                   //Initialize the used variable values
                   #temp32TempDword1 := 16#1;
                   #temp16IndexAnalog := 16#0;
                   #temp16IndexDigital := 16#0;
                   #temp16IndexBinary := 16#0;
                   #temp16IndexString := 16#0;
                   //Initialize the Procedure Para index and Name index while changing of Procedure and changing of screen selection b/w Prepared and Current procedure
                   IF ((#statLasProcedureCur <> #ProcedureCur) OR (#statLasProcedureReq <> #ProcedureReq) OR (#statLastReqProcedSelected <> #ProcedureParaType.ProcedureReqCurInd)) THEN
                       #ProcedureParaType.IndexAnalog := 16#0;
                       #ProcedureParaType.NameIndexAnalog := 16#0;
                       #ProcedureParaType.IndexDigital := 16#0;
                       #ProcedureParaType.NameIndexDigital := 16#0;
                       #ProcedureParaType.IndexBinary := 16#0;
                       #ProcedureParaType.NameIndexBinary := 16#0;
                       #ProcedureParaType.IndexString := 16#0;
                       #ProcedureParaType.NameIndexString := 16#0;
                   END_IF;
                   IF (((#ProcedureCur <> 16#0) AND NOT #ProcedureParaType.ProcedureReqCurInd) OR ((#ProcedureReq <> 16#0) AND #ProcedureParaType.ProcedureReqCurInd)) THEN
                       //Used/Mapped parameter count with individual parameter type will written from the Tool
                       #statTotalProcedureParameters := #MAPPED_PROCEDURE_ANALOG + #MAPPED_PROCEDURE_DIGITAL + #MAPPED_PROCEDURE_BINARY + #MAPPED_PROCEDURE_STRING - 1;
                       IF ((#statTotalProcedureParameters >= 0) AND (#statTotalProcedureParameters <= #PROCEDURE_PARAMETER_MAX)) THEN
                           FOR #temp16IndexOfDefinition := #PROCEDURE_PARAMETER_MIN TO #statTotalProcedureParameters BY 1 DO
                               // Condition for allow the loop iteration only within the start and end index
                               IF (((#stat16ProcParaEndIndex - #stat16ProcParaStartIndex) - #temp16IndexOfDefinition + #PROCEDURE_PARAMETER_MIN) >= 0) THEN
                                   #statInternalCurProcParameter[#temp16IndexOfDefinition].index := #tempSetup.stepOrder.parameterIndex[#stat16ProcParaStartIndex + #temp16IndexOfDefinition];  // MiS: content of first parameterIndex to first internal index, content of second parameterIndex to second internal index etc.
                                   #temp16Index := #statInternalCurProcParameter[#temp16IndexOfDefinition].index;//Move index info to the local var
                                   #temp16ParameterType := #tempSetup.step.parameterDefinition[#temp16Index].type;  // Get type of current parameter
                                   #temp16IndexMTP := #tempSetup.step.parameterDefinition[#temp16Index].indexMTP;//Get parameter indexMTP(wrapper DB) from the setup DB.
                                   #temp16IndexIO := #tempSetup.step.parameterDefinition[#temp16Index].indexIO;
                                   //Condition TO check parameter types are in the range
                                   IF (#temp16ParameterType >= #TYPE_NONE) AND (#temp16ParameterType <= #TYPE_STRING) THEN
                                       REGION Copy procedure parameters from input
                                           CASE #temp16ParameterType OF
                                                   // If Parameter type = 1(Analog)
                                               #TYPE_ANALOG:
                                                   REGION Analog
                                                       //Bit Masking funtionality for calculate the used Analog parameter and Position of the Parameter name in the HMI Text List                                              
                                                       #ProcedureParaType.IndexAnalog := #ProcedureParaType.IndexAnalog OR SHL(IN := #temp32TempDword1, N := INT_TO_UINT(#temp16IndexOfDefinition));
                                                       #ProcedureParaType.NameIndexAnalog := #ProcedureParaType.NameIndexAnalog OR SHL(IN := #temp32TempDword1, N := INT_TO_UINT(#temp16Index));
                                                       //WinCC Parameter View Faceplate logic
                                                       //#StatConfigPara.Analog[#temp16IndexIO] := #MTPConfigurationParameterAnalog[#temp16IndexMTP];
                                                       #ProcedureAna[#temp16IndexAnalog].WQC := #ProcedureParameterAnalog[#temp16IndexMTP].WQC;
                                                       #ProcedureAna[#temp16IndexAnalog].ApplyEn := #ProcedureParameterAnalog[#temp16IndexMTP].ApplyEn;
                                                       #ProcedureAna[#temp16IndexAnalog].ApplyInt := #ProcedureParameterAnalog[#temp16IndexMTP].ApplyInt;
                                                       #ProcedureAna[#temp16IndexAnalog].StateChannel := #ProcedureParameterAnalog[#temp16IndexMTP].StateChannel;
                                                       #ProcedureAna[#temp16IndexAnalog].StateOffAut := #ProcedureParameterAnalog[#temp16IndexMTP].StateOffAut;
                                                       #ProcedureAna[#temp16IndexAnalog].StateOpAut := #ProcedureParameterAnalog[#temp16IndexMTP].StateOpAut;
                                                       #ProcedureAna[#temp16IndexAnalog].StateAutAut := #ProcedureParameterAnalog[#temp16IndexMTP].StateAutAut;
                                                       #ProcedureAna[#temp16IndexAnalog].StateOffAct := #ProcedureParameterAnalog[#temp16IndexMTP].StateOffAct;
                                                       #ProcedureAna[#temp16IndexAnalog].StateOpAct := #ProcedureParameterAnalog[#temp16IndexMTP].StateOpAct;
                                                       #ProcedureAna[#temp16IndexAnalog].StateAutAct := #ProcedureParameterAnalog[#temp16IndexMTP].StateAutAct;
                                                       #ProcedureAna[#temp16IndexAnalog].SrcChannel := #ProcedureParameterAnalog[#temp16IndexMTP].SrcChannel;
                                                       #ProcedureAna[#temp16IndexAnalog].SrcExtAut := #ProcedureParameterAnalog[#temp16IndexMTP].SrcExtAut;
                                                       #ProcedureAna[#temp16IndexAnalog].SrcIntAut := #ProcedureParameterAnalog[#temp16IndexMTP].SrcIntAut;
                                                       #ProcedureAna[#temp16IndexAnalog].SrcIntAct := #ProcedureParameterAnalog[#temp16IndexMTP].SrcIntAct;
                                                       #ProcedureAna[#temp16IndexAnalog].SrcExtAct := #ProcedureParameterAnalog[#temp16IndexMTP].SrcExtAct;
                                                       #ProcedureAna[#temp16IndexAnalog].VInt := #ProcedureParameterAnalog[#temp16IndexMTP].VInt;
                                                       #ProcedureAna[#temp16IndexAnalog].VReq := #ProcedureParameterAnalog[#temp16IndexMTP].VReq;
                                                       #ProcedureAna[#temp16IndexAnalog].VOut := #ProcedureParameterAnalog[#temp16IndexMTP].VOut;
                                                       #ProcedureAna[#temp16IndexAnalog].VFbk := #ProcedureParameterAnalog[#temp16IndexMTP].VFbk;
                                                       #ProcedureAna[#temp16IndexAnalog].VSclMin := #ProcedureParameterAnalog[#temp16IndexMTP].VSclMin;
                                                       #ProcedureAna[#temp16IndexAnalog].VSclMax := #ProcedureParameterAnalog[#temp16IndexMTP].VSclMax;
                                                       #ProcedureAna[#temp16IndexAnalog].VUnit := #ProcedureParameterAnalog[#temp16IndexMTP].VUnit;
                                                       #ProcedureAna[#temp16IndexAnalog].VMin := #ProcedureParameterAnalog[#temp16IndexMTP].VMin;
                                                       #ProcedureAna[#temp16IndexAnalog].VMax := #ProcedureParameterAnalog[#temp16IndexMTP].VMax;
                                                       //Write values from WinCC
                                                       IF #ProcedureParameterAnalog[#temp16IndexMTP].OSLevel = #StatProcedureAnalog[#temp16IndexAnalog].OSLevel THEN
                                                           #ProcedureParameterAnalog[#temp16IndexMTP].OSLevel := #ProcedureAna[#temp16IndexAnalog].OSLevel;
                                                       ELSE
                                                           #ProcedureAna[#temp16IndexAnalog].OSLevel := #ProcedureParameterAnalog[#temp16IndexMTP].OSLevel;
                                                       END_IF;
                                                       IF #ProcedureParameterAnalog[#temp16IndexMTP].ApplyExt = #StatProcedureAnalog[#temp16IndexAnalog].ApplyExt THEN
                                                           #ProcedureParameterAnalog[#temp16IndexMTP].ApplyExt := #ProcedureAna[#temp16IndexAnalog].ApplyExt;
                                                       ELSE
                                                           #ProcedureAna[#temp16IndexAnalog].ApplyExt := #ProcedureParameterAnalog[#temp16IndexMTP].ApplyExt;
                                                       END_IF;
                                                       IF #ProcedureParameterAnalog[#temp16IndexMTP].ApplyOp = #StatProcedureAnalog[#temp16IndexAnalog].ApplyOp THEN
                                                           #ProcedureParameterAnalog[#temp16IndexMTP].ApplyOp := #ProcedureAna[#temp16IndexAnalog].ApplyOp;
                                                       ELSE
                                                           #ProcedureAna[#temp16IndexAnalog].ApplyOp := #ProcedureParameterAnalog[#temp16IndexMTP].ApplyOp;
                                                       END_IF;
                                                       IF #ProcedureParameterAnalog[#temp16IndexMTP].Sync = #StatProcedureAnalog[#temp16IndexAnalog].Sync THEN
                                                           #ProcedureParameterAnalog[#temp16IndexMTP].Sync := #ProcedureAna[#temp16IndexAnalog].Sync;
                                                       ELSE
                                                           #ProcedureAna[#temp16IndexAnalog].Sync := #ProcedureParameterAnalog[#temp16IndexMTP].Sync;
                                                       END_IF;
                                                       IF #ProcedureParameterAnalog[#temp16IndexMTP].StateOffOp = #StatProcedureAnalog[#temp16IndexAnalog].StateOffOp THEN
                                                           #ProcedureParameterAnalog[#temp16IndexMTP].StateOffOp := #ProcedureAna[#temp16IndexAnalog].StateOffOp;
                                                       ELSE
                                                           #ProcedureAna[#temp16IndexAnalog].StateOffOp := #ProcedureParameterAnalog[#temp16IndexMTP].StateOffOp;
                                                       END_IF;
                                                       IF #ProcedureParameterAnalog[#temp16IndexMTP].StateOpOp = #StatProcedureAnalog[#temp16IndexAnalog].StateOpOp THEN
                                                           #ProcedureParameterAnalog[#temp16IndexMTP].StateOpOp := #ProcedureAna[#temp16IndexAnalog].StateOpOp;
                                                       ELSE
                                                           #ProcedureAna[#temp16IndexAnalog].StateOpOp := #ProcedureParameterAnalog[#temp16IndexMTP].StateOpOp;
                                                       END_IF;
                                                       IF #ProcedureParameterAnalog[#temp16IndexMTP].StateAutOp = #StatProcedureAnalog[#temp16IndexAnalog].StateAutOp THEN
                                                           #ProcedureParameterAnalog[#temp16IndexMTP].StateAutOp := #ProcedureAna[#temp16IndexAnalog].StateAutOp;
                                                       ELSE
                                                           #ProcedureAna[#temp16IndexAnalog].StateAutOp := #ProcedureParameterAnalog[#temp16IndexMTP].StateAutOp;
                                                       END_IF;
                                                       IF #ProcedureParameterAnalog[#temp16IndexMTP].SrcIntOp = #StatProcedureAnalog[#temp16IndexAnalog].SrcIntOp THEN
                                                           #ProcedureParameterAnalog[#temp16IndexMTP].SrcIntOp := #ProcedureAna[#temp16IndexAnalog].SrcIntOp;
                                                       ELSE
                                                           #ProcedureAna[#temp16IndexAnalog].SrcIntOp := #ProcedureParameterAnalog[#temp16IndexMTP].SrcIntOp;
                                                       END_IF;
                                                       IF #ProcedureParameterAnalog[#temp16IndexMTP].SrcExtOp = #StatProcedureAnalog[#temp16IndexAnalog].SrcExtOp THEN
                                                           #ProcedureParameterAnalog[#temp16IndexMTP].SrcExtOp := #ProcedureAna[#temp16IndexAnalog].SrcExtOp;
                                                       ELSE
                                                           #ProcedureAna[#temp16IndexAnalog].SrcExtOp := #ProcedureParameterAnalog[#temp16IndexMTP].SrcExtOp;
                                                       END_IF;
                                                       IF #ProcedureParameterAnalog[#temp16IndexMTP].VExt = #StatProcedureAnalog[#temp16IndexAnalog].VExt THEN
                                                           #ProcedureParameterAnalog[#temp16IndexMTP].VExt := #ProcedureAna[#temp16IndexAnalog].VExt;
                                                       ELSE
                                                           #ProcedureAna[#temp16IndexAnalog].VExt := #ProcedureParameterAnalog[#temp16IndexMTP].VExt;
                                                       END_IF;
                                                       IF #ProcedureParameterAnalog[#temp16IndexMTP].VOp = #StatProcedureAnalog[#temp16IndexAnalog].VOp THEN
                                                           #ProcedureParameterAnalog[#temp16IndexMTP].VOp := #ProcedureAna[#temp16IndexAnalog].VOp;
                                                       ELSE
                                                           #ProcedureAna[#temp16IndexAnalog].VOp := #ProcedureParameterAnalog[#temp16IndexMTP].VOp;
                                                       END_IF;

                                                       #StatProcedureAnalog[#temp16IndexAnalog].OSLevel := #ProcedureAna[#temp16IndexAnalog].OSLevel;
                                                       #StatProcedureAnalog[#temp16IndexAnalog].ApplyExt := #ProcedureAna[#temp16IndexAnalog].ApplyExt;
                                                       #StatProcedureAnalog[#temp16IndexAnalog].ApplyOp := #ProcedureAna[#temp16IndexAnalog].ApplyOp;
                                                       #StatProcedureAnalog[#temp16IndexAnalog].Sync := #ProcedureAna[#temp16IndexAnalog].Sync;
                                                       #StatProcedureAnalog[#temp16IndexAnalog].StateOffOp := #ProcedureAna[#temp16IndexAnalog].StateOffOp;
                                                       #StatProcedureAnalog[#temp16IndexAnalog].StateOpOp := #ProcedureAna[#temp16IndexAnalog].StateOpOp;
                                                       #StatProcedureAnalog[#temp16IndexAnalog].StateAutOp := #ProcedureAna[#temp16IndexAnalog].StateAutOp;
                                                       #StatProcedureAnalog[#temp16IndexAnalog].SrcIntOp := #ProcedureAna[#temp16IndexAnalog].SrcIntOp;
                                                       #StatProcedureAnalog[#temp16IndexAnalog].SrcExtOp := #ProcedureAna[#temp16IndexAnalog].SrcExtOp;
                                                       #StatProcedureAnalog[#temp16IndexAnalog].VExt := #ProcedureAna[#temp16IndexAnalog].VExt;
                                                       #StatProcedureAnalog[#temp16IndexAnalog].VOp := #ProcedureAna[#temp16IndexAnalog].VOp;

                                                       #temp16IndexAnalog := #temp16IndexAnalog + 1;
                                                   END_REGION
                                                   // If Parameter type = 2(Digital)     
                                               #TYPE_DIGITAL:
                                                   REGION Digital
                                                       //Bit Masking funtionality for calculate the used Digital parameter and Position of the Parameter name in the HMI Text List  
                                                       #ProcedureParaType.IndexDigital := #ProcedureParaType.IndexDigital OR SHL(IN := #temp32TempDword1, N := INT_TO_UINT(#temp16IndexOfDefinition));
                                                       #ProcedureParaType.NameIndexDigital := #ProcedureParaType.NameIndexDigital OR SHL(IN := #temp32TempDword1, N := INT_TO_UINT(#temp16Index));
                                                       //WinCC Parameter View Faceplate logic
                                                       //#StatConfigPara.Digital[#temp16IndexIO] := #MTPConfigurationParameterAnalog[#temp16IndexMTP];
                                                       #ProcedureDint[#temp16IndexDigital].WQC := #ProcedureParameterDigital[#temp16IndexMTP].WQC;
                                                       #ProcedureDint[#temp16IndexDigital].ApplyEn := #ProcedureParameterDigital[#temp16IndexMTP].ApplyEn;
                                                       #ProcedureDint[#temp16IndexDigital].ApplyInt := #ProcedureParameterDigital[#temp16IndexMTP].ApplyInt;
                                                       #ProcedureDint[#temp16IndexDigital].StateChannel := #ProcedureParameterDigital[#temp16IndexMTP].StateChannel;
                                                       #ProcedureDint[#temp16IndexDigital].StateOffAut := #ProcedureParameterDigital[#temp16IndexMTP].StateOffAut;
                                                       #ProcedureDint[#temp16IndexDigital].StateOpAut := #ProcedureParameterDigital[#temp16IndexMTP].StateOpAut;
                                                       #ProcedureDint[#temp16IndexDigital].StateAutAut := #ProcedureParameterDigital[#temp16IndexMTP].StateAutAut;
                                                       #ProcedureDint[#temp16IndexDigital].StateOffAct := #ProcedureParameterDigital[#temp16IndexMTP].StateOffAct;
                                                       #ProcedureDint[#temp16IndexDigital].StateOpAct := #ProcedureParameterDigital[#temp16IndexMTP].StateOpAct;
                                                       #ProcedureDint[#temp16IndexDigital].StateAutAct := #ProcedureParameterDigital[#temp16IndexMTP].StateAutAct;
                                                       #ProcedureDint[#temp16IndexDigital].SrcChannel := #ProcedureParameterDigital[#temp16IndexMTP].SrcChannel;
                                                       #ProcedureDint[#temp16IndexDigital].SrcExtAut := #ProcedureParameterDigital[#temp16IndexMTP].SrcExtAut;
                                                       #ProcedureDint[#temp16IndexDigital].SrcIntAut := #ProcedureParameterDigital[#temp16IndexMTP].SrcIntAut;
                                                       #ProcedureDint[#temp16IndexDigital].SrcIntAct := #ProcedureParameterDigital[#temp16IndexMTP].SrcIntAct;
                                                       #ProcedureDint[#temp16IndexDigital].SrcExtAct := #ProcedureParameterDigital[#temp16IndexMTP].SrcExtAct;
                                                       #ProcedureDint[#temp16IndexDigital].VInt := #ProcedureParameterDigital[#temp16IndexMTP].VInt;
                                                       #ProcedureDint[#temp16IndexDigital].VReq := #ProcedureParameterDigital[#temp16IndexMTP].VReq;
                                                       #ProcedureDint[#temp16IndexDigital].VOut := #ProcedureParameterDigital[#temp16IndexMTP].VOut;
                                                       #ProcedureDint[#temp16IndexDigital].VFbk := #ProcedureParameterDigital[#temp16IndexMTP].VFbk;
                                                       #ProcedureDint[#temp16IndexDigital].VSclMin := #ProcedureParameterDigital[#temp16IndexMTP].VSclMin;
                                                       #ProcedureDint[#temp16IndexDigital].VSclMax := #ProcedureParameterDigital[#temp16IndexMTP].VSclMax;
                                                       #ProcedureDint[#temp16IndexDigital].VUnit := #ProcedureParameterDigital[#temp16IndexMTP].VUnit;
                                                       #ProcedureDint[#temp16IndexDigital].VMin := #ProcedureParameterDigital[#temp16IndexMTP].VMin;
                                                       #ProcedureDint[#temp16IndexDigital].VMax := #ProcedureParameterDigital[#temp16IndexMTP].VMax;
                                                       //Write values from WinCC
                                                       IF #ProcedureParameterDigital[#temp16IndexMTP].OSLevel = #StatProcedureDigital[#temp16IndexDigital].OSLevel THEN
                                                           #ProcedureParameterDigital[#temp16IndexMTP].OSLevel := #ProcedureDint[#temp16IndexDigital].OSLevel;
                                                       ELSE
                                                           #ProcedureDint[#temp16IndexDigital].OSLevel := #ProcedureParameterDigital[#temp16IndexMTP].OSLevel;
                                                       END_IF;
                                                       IF #ProcedureParameterDigital[#temp16IndexMTP].ApplyExt = #StatProcedureDigital[#temp16IndexDigital].ApplyExt THEN
                                                           #ProcedureParameterDigital[#temp16IndexMTP].ApplyExt := #ProcedureDint[#temp16IndexDigital].ApplyExt;
                                                       ELSE
                                                           #ProcedureDint[#temp16IndexDigital].ApplyExt := #ProcedureParameterDigital[#temp16IndexMTP].ApplyExt;
                                                       END_IF;
                                                       IF #ProcedureParameterDigital[#temp16IndexMTP].ApplyOp = #StatProcedureDigital[#temp16IndexDigital].ApplyOp THEN
                                                           #ProcedureParameterDigital[#temp16IndexMTP].ApplyOp := #ProcedureDint[#temp16IndexDigital].ApplyOp;
                                                       ELSE
                                                           #ProcedureDint[#temp16IndexDigital].ApplyOp := #ProcedureParameterDigital[#temp16IndexMTP].ApplyOp;
                                                       END_IF;
                                                       IF #ProcedureParameterDigital[#temp16IndexMTP].Sync = #StatProcedureDigital[#temp16IndexDigital].Sync THEN
                                                           #ProcedureParameterDigital[#temp16IndexMTP].Sync := #ProcedureDint[#temp16IndexDigital].Sync;
                                                       ELSE
                                                           #ProcedureDint[#temp16IndexDigital].Sync := #ProcedureParameterDigital[#temp16IndexMTP].Sync;
                                                       END_IF;
                                                       IF #ProcedureParameterDigital[#temp16IndexMTP].StateOffOp = #StatProcedureDigital[#temp16IndexDigital].StateOffOp THEN
                                                           #ProcedureParameterDigital[#temp16IndexMTP].StateOffOp := #ProcedureDint[#temp16IndexDigital].StateOffOp;
                                                       ELSE
                                                           #ProcedureDint[#temp16IndexDigital].StateOffOp := #ProcedureParameterDigital[#temp16IndexMTP].StateOffOp;
                                                       END_IF;
                                                       IF #ProcedureParameterDigital[#temp16IndexMTP].StateOpOp = #StatProcedureDigital[#temp16IndexDigital].StateOpOp THEN
                                                           #ProcedureParameterDigital[#temp16IndexMTP].StateOpOp := #ProcedureDint[#temp16IndexDigital].StateOpOp;
                                                       ELSE
                                                           #ProcedureDint[#temp16IndexDigital].StateOpOp := #ProcedureParameterDigital[#temp16IndexMTP].StateOpOp;
                                                       END_IF;
                                                       IF #ProcedureParameterDigital[#temp16IndexMTP].StateAutOp = #StatProcedureDigital[#temp16IndexDigital].StateAutOp THEN
                                                           #ProcedureParameterDigital[#temp16IndexMTP].StateAutOp := #ProcedureDint[#temp16IndexDigital].StateAutOp;
                                                       ELSE
                                                           #ProcedureDint[#temp16IndexDigital].StateAutOp := #ProcedureParameterDigital[#temp16IndexMTP].StateAutOp;
                                                       END_IF;
                                                       IF #ProcedureParameterDigital[#temp16IndexMTP].SrcIntOp = #StatProcedureDigital[#temp16IndexDigital].SrcIntOp THEN
                                                           #ProcedureParameterDigital[#temp16IndexMTP].SrcIntOp := #ProcedureDint[#temp16IndexDigital].SrcIntOp;
                                                       ELSE
                                                           #ProcedureDint[#temp16IndexDigital].SrcIntOp := #ProcedureParameterDigital[#temp16IndexMTP].SrcIntOp;
                                                       END_IF;
                                                       IF #ProcedureParameterDigital[#temp16IndexMTP].SrcExtOp = #StatProcedureDigital[#temp16IndexDigital].SrcExtOp THEN
                                                           #ProcedureParameterDigital[#temp16IndexMTP].SrcExtOp := #ProcedureDint[#temp16IndexDigital].SrcExtOp;
                                                       ELSE
                                                           #ProcedureDint[#temp16IndexDigital].SrcExtOp := #ProcedureParameterDigital[#temp16IndexMTP].SrcExtOp;
                                                       END_IF;
                                                       IF #ProcedureParameterDigital[#temp16IndexMTP].VExt = #StatProcedureDigital[#temp16IndexDigital].VExt THEN
                                                           #ProcedureParameterDigital[#temp16IndexMTP].VExt := #ProcedureDint[#temp16IndexDigital].VExt;
                                                       ELSE
                                                           #ProcedureDint[#temp16IndexDigital].VExt := #ProcedureParameterDigital[#temp16IndexMTP].VExt;
                                                       END_IF;
                                                       IF #ProcedureParameterDigital[#temp16IndexMTP].VOp = #StatProcedureDigital[#temp16IndexDigital].VOp THEN
                                                           #ProcedureParameterDigital[#temp16IndexMTP].VOp := #ProcedureDint[#temp16IndexDigital].VOp;
                                                       ELSE
                                                           #ProcedureDint[#temp16IndexDigital].VOp := #ProcedureParameterDigital[#temp16IndexMTP].VOp;
                                                       END_IF;

                                                       #StatProcedureDigital[#temp16IndexDigital].OSLevel := #ProcedureDint[#temp16IndexDigital].OSLevel;
                                                       #StatProcedureDigital[#temp16IndexDigital].ApplyExt := #ProcedureDint[#temp16IndexDigital].ApplyExt;
                                                       #StatProcedureDigital[#temp16IndexDigital].ApplyOp := #ProcedureDint[#temp16IndexDigital].ApplyOp;
                                                       #StatProcedureDigital[#temp16IndexDigital].Sync := #ProcedureDint[#temp16IndexDigital].Sync;
                                                       #StatProcedureDigital[#temp16IndexDigital].StateOffOp := #ProcedureDint[#temp16IndexDigital].StateOffOp;
                                                       #StatProcedureDigital[#temp16IndexDigital].StateOpOp := #ProcedureDint[#temp16IndexDigital].StateOpOp;
                                                       #StatProcedureDigital[#temp16IndexDigital].StateAutOp := #ProcedureDint[#temp16IndexDigital].StateAutOp;
                                                       #StatProcedureDigital[#temp16IndexDigital].SrcIntOp := #ProcedureDint[#temp16IndexDigital].SrcIntOp;
                                                       #StatProcedureDigital[#temp16IndexDigital].SrcExtOp := #ProcedureDint[#temp16IndexDigital].SrcExtOp;
                                                       #StatProcedureDigital[#temp16IndexDigital].VExt := #ProcedureDint[#temp16IndexDigital].VExt;
                                                       #StatProcedureDigital[#temp16IndexDigital].VOp := #ProcedureDint[#temp16IndexDigital].VOp;

                                                       #temp16IndexDigital := #temp16IndexDigital + 1;
                                                   END_REGION
                                                   // If Parameter type = 3(Binary)    
                                               #TYPE_BINARY:
                                                   REGION Binary
                                                       //Bit Masking funtionality for calculate the used Binary parameter and Position of the Parameter name in the HMI Text List  
                                                       #ProcedureParaType.IndexBinary := #ProcedureParaType.IndexBinary OR SHL(IN := #temp32TempDword1, N := INT_TO_UINT(#temp16IndexOfDefinition));
                                                       #ProcedureParaType.NameIndexBinary := #ProcedureParaType.NameIndexBinary OR SHL(IN := #temp32TempDword1, N := INT_TO_UINT(#temp16Index));
                                                       //WinCC Parameter View Faceplate logic
                                                       //#StatConfigPara.Binary[#temp16IndexIO] := #MTPConfigurationParameterAnalog[#temp16IndexMTP];
                                                       #ProcedureBin[#temp16IndexBinary].WQC := #ProcedureParameterBinary[#temp16IndexMTP].WQC;
                                                       #ProcedureBin[#temp16IndexBinary].ApplyEn := #ProcedureParameterBinary[#temp16IndexMTP].ApplyEn;
                                                       #ProcedureBin[#temp16IndexBinary].ApplyInt := #ProcedureParameterBinary[#temp16IndexMTP].ApplyInt;
                                                       #ProcedureBin[#temp16IndexBinary].StateChannel := #ProcedureParameterBinary[#temp16IndexMTP].StateChannel;
                                                       #ProcedureBin[#temp16IndexBinary].StateOffAut := #ProcedureParameterBinary[#temp16IndexMTP].StateOffAut;
                                                       #ProcedureBin[#temp16IndexBinary].StateOpAut := #ProcedureParameterBinary[#temp16IndexMTP].StateOpAut;
                                                       #ProcedureBin[#temp16IndexBinary].StateAutAut := #ProcedureParameterBinary[#temp16IndexMTP].StateAutAut;
                                                       #ProcedureBin[#temp16IndexBinary].StateOffAct := #ProcedureParameterBinary[#temp16IndexMTP].StateOffAct;
                                                       #ProcedureBin[#temp16IndexBinary].StateOpAct := #ProcedureParameterBinary[#temp16IndexMTP].StateOpAct;
                                                       #ProcedureBin[#temp16IndexBinary].StateAutAct := #ProcedureParameterBinary[#temp16IndexMTP].StateAutAct;
                                                       #ProcedureBin[#temp16IndexBinary].SrcChannel := #ProcedureParameterBinary[#temp16IndexMTP].SrcChannel;
                                                       #ProcedureBin[#temp16IndexBinary].SrcExtAut := #ProcedureParameterBinary[#temp16IndexMTP].SrcExtAut;
                                                       #ProcedureBin[#temp16IndexBinary].SrcIntAut := #ProcedureParameterBinary[#temp16IndexMTP].SrcIntAut;
                                                       #ProcedureBin[#temp16IndexBinary].SrcIntAct := #ProcedureParameterBinary[#temp16IndexMTP].SrcIntAct;
                                                       #ProcedureBin[#temp16IndexBinary].SrcExtAct := #ProcedureParameterBinary[#temp16IndexMTP].SrcExtAct;
                                                       #ProcedureBin[#temp16IndexBinary].VInt := #ProcedureParameterBinary[#temp16IndexMTP].VInt;
                                                       #ProcedureBin[#temp16IndexBinary].VReq := #ProcedureParameterBinary[#temp16IndexMTP].VReq;
                                                       #ProcedureBin[#temp16IndexBinary].VOut := #ProcedureParameterBinary[#temp16IndexMTP].VOut;
                                                       #ProcedureBin[#temp16IndexBinary].VFbk := #ProcedureParameterBinary[#temp16IndexMTP].VFbk;

                                                       //Write values from WinCC
                                                       IF #ProcedureParameterBinary[#temp16IndexMTP].OSLevel = #StatProcedureBinary[#temp16IndexBinary].OSLevel THEN
                                                           #ProcedureParameterBinary[#temp16IndexMTP].OSLevel := #ProcedureBin[#temp16IndexBinary].OSLevel;
                                                       ELSE
                                                           #ProcedureBin[#temp16IndexBinary].OSLevel := #ProcedureParameterBinary[#temp16IndexMTP].OSLevel;
                                                       END_IF;
                                                       IF #ProcedureParameterBinary[#temp16IndexMTP].ApplyExt = #StatProcedureBinary[#temp16IndexBinary].ApplyExt THEN
                                                           #ProcedureParameterBinary[#temp16IndexMTP].ApplyExt := #ProcedureBin[#temp16IndexBinary].ApplyExt;
                                                       ELSE
                                                           #ProcedureBin[#temp16IndexBinary].ApplyExt := #ProcedureParameterBinary[#temp16IndexMTP].ApplyExt;
                                                       END_IF;
                                                       IF #ProcedureParameterBinary[#temp16IndexMTP].ApplyOp = #StatProcedureBinary[#temp16IndexBinary].ApplyOp THEN
                                                           #ProcedureParameterBinary[#temp16IndexMTP].ApplyOp := #ProcedureBin[#temp16IndexBinary].ApplyOp;
                                                       ELSE
                                                           #ProcedureBin[#temp16IndexBinary].ApplyOp := #ProcedureParameterBinary[#temp16IndexMTP].ApplyOp;
                                                       END_IF;
                                                       IF #ProcedureParameterBinary[#temp16IndexMTP].Sync = #StatProcedureBinary[#temp16IndexBinary].Sync THEN
                                                           #ProcedureParameterBinary[#temp16IndexMTP].Sync := #ProcedureBin[#temp16IndexBinary].Sync;
                                                       ELSE
                                                           #ProcedureBin[#temp16IndexBinary].Sync := #ProcedureParameterBinary[#temp16IndexMTP].Sync;
                                                       END_IF;
                                                       IF #ProcedureParameterBinary[#temp16IndexMTP].StateOffOp = #StatProcedureBinary[#temp16IndexBinary].StateOffOp THEN
                                                           #ProcedureParameterBinary[#temp16IndexMTP].StateOffOp := #ProcedureBin[#temp16IndexBinary].StateOffOp;
                                                       ELSE
                                                           #ProcedureBin[#temp16IndexBinary].StateOffOp := #ProcedureParameterBinary[#temp16IndexMTP].StateOffOp;
                                                       END_IF;
                                                       IF #ProcedureParameterBinary[#temp16IndexMTP].StateOpOp = #StatProcedureBinary[#temp16IndexBinary].StateOpOp THEN
                                                           #ProcedureParameterBinary[#temp16IndexMTP].StateOpOp := #ProcedureBin[#temp16IndexBinary].StateOpOp;
                                                       ELSE
                                                           #ProcedureBin[#temp16IndexBinary].StateOpOp := #ProcedureParameterBinary[#temp16IndexMTP].StateOpOp;
                                                       END_IF;
                                                       IF #ProcedureParameterBinary[#temp16IndexMTP].StateAutOp = #StatProcedureBinary[#temp16IndexBinary].StateAutOp THEN
                                                           #ProcedureParameterBinary[#temp16IndexMTP].StateAutOp := #ProcedureBin[#temp16IndexBinary].StateAutOp;
                                                       ELSE
                                                           #ProcedureBin[#temp16IndexBinary].StateAutOp := #ProcedureParameterBinary[#temp16IndexMTP].StateAutOp;
                                                       END_IF;
                                                       IF #ProcedureParameterBinary[#temp16IndexMTP].SrcIntOp = #StatProcedureBinary[#temp16IndexBinary].SrcIntOp THEN
                                                           #ProcedureParameterBinary[#temp16IndexMTP].SrcIntOp := #ProcedureBin[#temp16IndexBinary].SrcIntOp;
                                                       ELSE
                                                           #ProcedureBin[#temp16IndexBinary].SrcIntOp := #ProcedureParameterBinary[#temp16IndexMTP].SrcIntOp;
                                                       END_IF;
                                                       IF #ProcedureParameterBinary[#temp16IndexMTP].SrcExtOp = #StatProcedureBinary[#temp16IndexBinary].SrcExtOp THEN
                                                           #ProcedureParameterBinary[#temp16IndexMTP].SrcExtOp := #ProcedureBin[#temp16IndexBinary].SrcExtOp;
                                                       ELSE
                                                           #ProcedureBin[#temp16IndexBinary].SrcExtOp := #ProcedureParameterBinary[#temp16IndexMTP].SrcExtOp;
                                                       END_IF;
                                                       IF #ProcedureParameterBinary[#temp16IndexMTP].VExt = #StatProcedureBinary[#temp16IndexBinary].VExt THEN
                                                           #ProcedureParameterBinary[#temp16IndexMTP].VExt := #ProcedureBin[#temp16IndexBinary].VExt;
                                                       ELSE
                                                           #ProcedureBin[#temp16IndexBinary].VExt := #ProcedureParameterBinary[#temp16IndexMTP].VExt;
                                                       END_IF;
                                                       IF #ProcedureParameterBinary[#temp16IndexMTP].VOp = #StatProcedureBinary[#temp16IndexBinary].VOp THEN
                                                           #ProcedureParameterBinary[#temp16IndexMTP].VOp := #ProcedureBin[#temp16IndexBinary].VOp;
                                                       ELSE
                                                           #ProcedureBin[#temp16IndexBinary].VOp := #ProcedureParameterBinary[#temp16IndexMTP].VOp;
                                                       END_IF;

                                                       #StatProcedureBinary[#temp16IndexBinary].OSLevel := #ProcedureBin[#temp16IndexBinary].OSLevel;
                                                       #StatProcedureBinary[#temp16IndexBinary].ApplyExt := #ProcedureBin[#temp16IndexBinary].ApplyExt;
                                                       #StatProcedureBinary[#temp16IndexBinary].ApplyOp := #ProcedureBin[#temp16IndexBinary].ApplyOp;
                                                       #StatProcedureBinary[#temp16IndexBinary].Sync := #ProcedureBin[#temp16IndexBinary].Sync;
                                                       #StatProcedureBinary[#temp16IndexBinary].StateOffOp := #ProcedureBin[#temp16IndexBinary].StateOffOp;
                                                       #StatProcedureBinary[#temp16IndexBinary].StateOpOp := #ProcedureBin[#temp16IndexBinary].StateOpOp;
                                                       #StatProcedureBinary[#temp16IndexBinary].StateAutOp := #ProcedureBin[#temp16IndexBinary].StateAutOp;
                                                       #StatProcedureBinary[#temp16IndexBinary].SrcIntOp := #ProcedureBin[#temp16IndexBinary].SrcIntOp;
                                                       #StatProcedureBinary[#temp16IndexBinary].SrcExtOp := #ProcedureBin[#temp16IndexBinary].SrcExtOp;
                                                       #StatProcedureBinary[#temp16IndexBinary].VExt := #ProcedureBin[#temp16IndexBinary].VExt;
                                                       #StatProcedureBinary[#temp16IndexBinary].VOp := #ProcedureBin[#temp16IndexBinary].VOp;

                                                       #temp16IndexBinary := #temp16IndexBinary + 1;
                                                   END_REGION
                                                   // If Parameter type = 4(String)    
                                               #TYPE_STRING:
                                                   REGION String
                                                       //Bit Masking funtionality for calculate the used String parameter and Position of the Parameter name in the HMI Text List  
                                                       #ProcedureParaType.IndexString := #ProcedureParaType.IndexString OR SHL(IN := #temp32TempDword1, N := INT_TO_UINT(#temp16IndexOfDefinition));
                                                       #ProcedureParaType.NameIndexString := #ProcedureParaType.NameIndexString OR SHL(IN := #temp32TempDword1, N := INT_TO_UINT(#temp16Index));
                                                       //WinCC Parameter View Faceplate logic
                                                       //#StatConfigPara."String"[#temp16IndexIO] := #MTPConfigurationParameterString[#temp16IndexMTP];
                                                       #ProcedureString[#temp16IndexString].WQC := #ProcedureParameterString[#temp16IndexMTP].WQC;
                                                       #ProcedureString[#temp16IndexString].ApplyEn := #ProcedureParameterString[#temp16IndexMTP].ApplyEn;
                                                       #ProcedureString[#temp16IndexString].ApplyInt := #ProcedureParameterString[#temp16IndexMTP].ApplyInt;
                                                       #ProcedureString[#temp16IndexString].StateChannel := #ProcedureParameterString[#temp16IndexMTP].StateChannel;
                                                       #ProcedureString[#temp16IndexString].StateOffAut := #ProcedureParameterString[#temp16IndexMTP].StateOffAut;
                                                       #ProcedureString[#temp16IndexString].StateOpAut := #ProcedureParameterString[#temp16IndexMTP].StateOpAut;
                                                       #ProcedureString[#temp16IndexString].StateAutAut := #ProcedureParameterString[#temp16IndexMTP].StateAutAut;
                                                       #ProcedureString[#temp16IndexString].StateOffAct := #ProcedureParameterString[#temp16IndexMTP].StateOffAct;
                                                       #ProcedureString[#temp16IndexString].StateOpAct := #ProcedureParameterString[#temp16IndexMTP].StateOpAct;
                                                       #ProcedureString[#temp16IndexString].StateAutAct := #ProcedureParameterString[#temp16IndexMTP].StateAutAct;
                                                       #ProcedureString[#temp16IndexString].SrcChannel := #ProcedureParameterString[#temp16IndexMTP].SrcChannel;
                                                       #ProcedureString[#temp16IndexString].SrcExtAut := #ProcedureParameterString[#temp16IndexMTP].SrcExtAut;
                                                       #ProcedureString[#temp16IndexString].SrcIntAut := #ProcedureParameterString[#temp16IndexMTP].SrcIntAut;
                                                       #ProcedureString[#temp16IndexString].SrcIntAct := #ProcedureParameterString[#temp16IndexMTP].SrcIntAct;
                                                       #ProcedureString[#temp16IndexString].SrcExtAct := #ProcedureParameterString[#temp16IndexMTP].SrcExtAct;
                                                       #ProcedureString[#temp16IndexString].VInt := #ProcedureParameterString[#temp16IndexMTP].VInt;
                                                       #ProcedureString[#temp16IndexString].VReq := #ProcedureParameterString[#temp16IndexMTP].VReq;
                                                       #ProcedureString[#temp16IndexString].VOut := #ProcedureParameterString[#temp16IndexMTP].VOut;
                                                       #ProcedureString[#temp16IndexString].VFbk := #ProcedureParameterString[#temp16IndexMTP].VFbk;

                                                       //Write values from WinCC
                                                       IF #ProcedureParameterString[#temp16IndexMTP].OSLevel = #StatProcedureString[#temp16IndexString].OSLevel THEN
                                                           #ProcedureParameterString[#temp16IndexMTP].OSLevel := #ProcedureString[#temp16IndexString].OSLevel;
                                                       ELSE
                                                           #ProcedureString[#temp16IndexString].OSLevel := #ProcedureParameterString[#temp16IndexMTP].OSLevel;
                                                       END_IF;
                                                       IF #ProcedureParameterString[#temp16IndexMTP].ApplyExt = #StatProcedureString[#temp16IndexString].ApplyExt THEN
                                                           #ProcedureParameterString[#temp16IndexMTP].ApplyExt := #ProcedureString[#temp16IndexString].ApplyExt;
                                                       ELSE
                                                           #ProcedureString[#temp16IndexString].ApplyExt := #ProcedureParameterString[#temp16IndexMTP].ApplyExt;
                                                       END_IF;
                                                       IF #ProcedureParameterString[#temp16IndexMTP].ApplyOp = #StatProcedureString[#temp16IndexString].ApplyOp THEN
                                                           #ProcedureParameterString[#temp16IndexMTP].ApplyOp := #ProcedureString[#temp16IndexString].ApplyOp;
                                                       ELSE
                                                           #ProcedureString[#temp16IndexString].ApplyOp := #ProcedureParameterString[#temp16IndexMTP].ApplyOp;
                                                       END_IF;
                                                       IF #ProcedureParameterString[#temp16IndexMTP].Sync = #StatProcedureString[#temp16IndexString].Sync THEN
                                                           #ProcedureParameterString[#temp16IndexMTP].Sync := #ProcedureString[#temp16IndexString].Sync;
                                                       ELSE
                                                           #ProcedureString[#temp16IndexString].Sync := #ProcedureParameterString[#temp16IndexMTP].Sync;
                                                       END_IF;
                                                       IF #ProcedureParameterString[#temp16IndexMTP].StateOffOp = #StatProcedureString[#temp16IndexString].StateOffOp THEN
                                                           #ProcedureParameterString[#temp16IndexMTP].StateOffOp := #ProcedureString[#temp16IndexString].StateOffOp;
                                                       ELSE
                                                           #ProcedureString[#temp16IndexString].StateOffOp := #ProcedureParameterString[#temp16IndexMTP].StateOffOp;
                                                       END_IF;
                                                       IF #ProcedureParameterString[#temp16IndexMTP].StateOpOp = #StatProcedureString[#temp16IndexString].StateOpOp THEN
                                                           #ProcedureParameterString[#temp16IndexMTP].StateOpOp := #ProcedureString[#temp16IndexString].StateOpOp;
                                                       ELSE
                                                           #ProcedureString[#temp16IndexString].StateOpOp := #ProcedureParameterString[#temp16IndexMTP].StateOpOp;
                                                       END_IF;
                                                       IF #ProcedureParameterString[#temp16IndexMTP].StateAutOp = #StatProcedureString[#temp16IndexString].StateAutOp THEN
                                                           #ProcedureParameterString[#temp16IndexMTP].StateAutOp := #ProcedureString[#temp16IndexString].StateAutOp;
                                                       ELSE
                                                           #ProcedureString[#temp16IndexString].StateAutOp := #ProcedureParameterString[#temp16IndexMTP].StateAutOp;
                                                       END_IF;
                                                       IF #ProcedureParameterString[#temp16IndexMTP].SrcIntOp = #StatProcedureString[#temp16IndexString].SrcIntOp THEN
                                                           #ProcedureParameterString[#temp16IndexMTP].SrcIntOp := #ProcedureString[#temp16IndexString].SrcIntOp;
                                                       ELSE
                                                           #ProcedureString[#temp16IndexString].SrcIntOp := #ProcedureParameterString[#temp16IndexMTP].SrcIntOp;
                                                       END_IF;
                                                       IF #ProcedureParameterString[#temp16IndexMTP].SrcExtOp = #StatProcedureString[#temp16IndexString].SrcExtOp THEN
                                                           #ProcedureParameterString[#temp16IndexMTP].SrcExtOp := #ProcedureString[#temp16IndexString].SrcExtOp;
                                                       ELSE
                                                           #ProcedureString[#temp16IndexString].SrcExtOp := #ProcedureParameterString[#temp16IndexMTP].SrcExtOp;
                                                       END_IF;
                                                       IF #ProcedureParameterString[#temp16IndexMTP].VExt = #StatProcedureString[#temp16IndexString].VExt THEN
                                                           #ProcedureParameterString[#temp16IndexMTP].VExt := #ProcedureString[#temp16IndexString].VExt;
                                                       ELSE
                                                           #ProcedureString[#temp16IndexString].VExt := #ProcedureParameterString[#temp16IndexMTP].VExt;
                                                       END_IF;
                                                       IF #ProcedureParameterString[#temp16IndexMTP].VOp = #StatProcedureString[#temp16IndexString].VOp THEN
                                                           #ProcedureParameterString[#temp16IndexMTP].VOp := #ProcedureString[#temp16IndexString].VOp;
                                                       ELSE
                                                           #ProcedureString[#temp16IndexString].VOp := #ProcedureParameterString[#temp16IndexMTP].VOp;
                                                       END_IF;

                                                       #StatProcedureString[#temp16IndexString].OSLevel := #ProcedureString[#temp16IndexString].OSLevel;
                                                       #StatProcedureString[#temp16IndexString].ApplyExt := #ProcedureString[#temp16IndexString].ApplyExt;
                                                       #StatProcedureString[#temp16IndexString].ApplyOp := #ProcedureString[#temp16IndexString].ApplyOp;
                                                       #StatProcedureString[#temp16IndexString].Sync := #ProcedureString[#temp16IndexString].Sync;
                                                       #StatProcedureString[#temp16IndexString].StateOffOp := #ProcedureString[#temp16IndexString].StateOffOp;
                                                       #StatProcedureString[#temp16IndexString].StateOpOp := #ProcedureString[#temp16IndexString].StateOpOp;
                                                       #StatProcedureString[#temp16IndexString].StateAutOp := #ProcedureString[#temp16IndexString].StateAutOp;
                                                       #StatProcedureString[#temp16IndexString].SrcIntOp := #ProcedureString[#temp16IndexString].SrcIntOp;
                                                       #StatProcedureString[#temp16IndexString].SrcExtOp := #ProcedureString[#temp16IndexString].SrcExtOp;
                                                       #StatProcedureString[#temp16IndexString].VExt := #ProcedureString[#temp16IndexString].VExt;
                                                       #StatProcedureString[#temp16IndexString].VOp := #ProcedureString[#temp16IndexString].VOp;

                                                       #temp16IndexString := #temp16IndexString + 1;
                                                   END_REGION
                                           END_CASE;
                                       END_REGION
                                   END_IF;
                               END_IF;
                           END_FOR;
                       END_IF;
                   END_IF;
               END_IF;
           END_REGION
       END_REGION

       REGION Process In Values

           REGION Get Start and End index details of the Current /Prepared procedure
               //Current/Prepared procedure selection for parameter display in the faceplate
               //#stat32PrecedureProcessInMap := -1;
               IF NOT (#ProcessInValueType.ProcedureReqCurInd) THEN
                   #stat32PrecedureProcessInMap := #tempSetup.procedure.procedure[#stat16ProceCurIndex].ProcedureProcessInMap[0];
               ELSIF (#ProcessInValueType.ProcedureReqCurInd) THEN
                   #stat32PrecedureProcessInMap := #tempSetup.procedure.procedure[#stat16ProceReqIndex].ProcedureProcessInMap[0];
               END_IF;
           END_REGION
           //Initialize the used variable values        
           #temp32TempDword1 := 16#1;
           #temp16IndexAnalog := 16#0;
           #temp16IndexDigital := 16#0;
           #temp16IndexBinary := 16#0;
           #temp16IndexString := 16#0;
           //Initialize the Process In Value index and Name index while changing of Procedure and changing of screen selection b/w Prepared and Current procedure
           IF ((#statLasProcedureCur <> #ProcedureCur) OR (#statLasProcedureReq <> #ProcedureReq) OR (#StatLastProceselProcessIn <> #ProcessInValueType.ProcedureReqCurInd)
               OR (((#ProcedureCur = 16#0) AND NOT #ProcessInValueType.ProcedureReqCurInd) OR ((#ProcedureReq = 16#0) AND #ProcessInValueType.ProcedureReqCurInd))) THEN
               #ProcessInValueType.IndexAnalog := 16#0;
               #ProcessInValueType.NameIndexAnalog := 16#0;
               #ProcessInValueType.IndexDigital := 16#0;
               #ProcessInValueType.NameIndexDigital := 16#0;
               #ProcessInValueType.IndexBinary := 16#0;
               #ProcessInValueType.NameIndexBinary := 16#0;
               #ProcessInValueType.IndexString := 16#0;
               #ProcessInValueType.NameIndexString := 16#0;
           END_IF;
           //Used/Mapped parameter count with individual parameter type will written from the Tool
           #statTotalProcessInValues := #MAPPED_PROCESS_IN_ANALOG + #MAPPED_PROCESS_IN_DIGITAL + #MAPPED_PROCESS_IN_BINARY + #MAPPED_PROCESS_IN_STRING - 1;
           IF (((#ProcedureCur <> 16#0) AND NOT #ProcessInValueType.ProcedureReqCurInd) OR ((#ProcedureReq <> 16#0) AND #ProcessInValueType.ProcedureReqCurInd)) THEN
               IF ((#statTotalProcessInValues >= 0) AND (#statTotalProcessInValues <= #PROCESS_VALUES_IN_MAX)) THEN
                   #temp16IndexOfDefinitionProcessIn := 16#0;
                   FOR #temp16IndexOfDefinition := #PROCESS_VALUES_IN_MIN TO #statTotalProcessInValues BY 1 DO
                       #temp16ParameterCMAddress := BYTE_TO_INT(#tempSetup.processValueInData.definition[#temp16IndexOfDefinition].controlModule);
                       #temp16ParameterType := #tempSetup.processValueInData.definition[#temp16IndexOfDefinition].type;
                       #temp16IndexMTP := #tempSetup.processValueInData.definition[#temp16IndexOfDefinition].indexMTP;
                       #tempUsed := #tempSetup.processValueInData.used;
                       // Find the procedure information assigned with the processIn values
                       IF (((#stat32PrecedureProcessInMap AND SHL(IN := #temp32TempDword1, N := INT_TO_UINT(#temp16IndexOfDefinition))) <> 0) = TRUE) THEN
                           #temp16IndexIO := #tempSetup.processValueInData.definition[#temp16IndexOfDefinition].indexIO;

                           IF (#temp16ParameterCMAddress <> 255) AND (#temp16ParameterCMAddress >= #NUMBER_OF_CONTROLMODULES_MIN) AND (#temp16ParameterCMAddress <= #NUMBER_OF_CONTROLMODULES)
                               AND (#temp16ParameterType >= #TYPE_NONE) AND (#temp16ParameterType <= #TYPE_STRING) THEN
                               #temp16TempInt1 := #temp16ParameterCMAddress / 32;    //DWORD - Adress
                               #temp16TempInt2 := #temp16ParameterCMAddress MOD 32;  //Bit - Adress
                               //If parameter is forced (FRC) --> Parameter is used
                               IF (((#tempUsed[#temp16TempInt1] AND SHL(IN := #temp32TempDword1, N := INT_TO_UINT(#temp16TempInt2))) <> 0) = TRUE) THEN
                                   CASE #temp16ParameterType OF
                                           // Check of mode is done in satellite blocks
                                       #TYPE_ANALOG:
                                           REGION Analog
                                               //Bit Masking funtionality for calculate the used Analog parameter and Position of the Parameter name in the HMI Text List 
                                               #ProcessInValueType.IndexAnalog := #ProcessInValueType.IndexAnalog OR SHL(IN := #temp32TempDword1, N := INT_TO_UINT(#temp16IndexOfDefinitionProcessIn));
                                               #ProcessInValueType.NameIndexAnalog := #ProcessInValueType.NameIndexAnalog OR SHL(IN := #temp32TempDword1, N := INT_TO_UINT(#temp16IndexOfDefinition));
                                               IF ((#temp16IndexIO >= #PROCESS_VALUES_IN_MIN) AND (#temp16IndexIO <= #PROCESS_VALUES_IN_ANALOG_MAX)) THEN
                                                   //WinCC Parameter View Faceplate logic
                                                   #ProcessInAna[#temp16IndexAnalog].WQC := #ProcessValueInAnalog[#temp16IndexMTP].WQC;
                                                   #ProcessInAna[#temp16IndexAnalog].OSLevel := #ProcessValueInAnalog[#temp16IndexMTP].OSLevel;
                                                   #ProcessInAna[#temp16IndexAnalog].V := #ProcessValueInAnalog[#temp16IndexMTP].V;
                                                   #ProcessInAna[#temp16IndexAnalog].VQC := #ProcessValueInAnalog[#temp16IndexMTP].VQC;
                                                   #ProcessInAna[#temp16IndexAnalog].SclMinCur := #ProcessValueInAnalog[#temp16IndexMTP].SclMinCur;
                                                   #ProcessInAna[#temp16IndexAnalog].SclMaxCur := #ProcessValueInAnalog[#temp16IndexMTP].SclMaxCur;
                                                   #ProcessInAna[#temp16IndexAnalog].UnitCur := #ProcessValueInAnalog[#temp16IndexMTP].UnitCur;
                                                   #ProcessInAna[#temp16IndexAnalog].SclMinExt := #ProcessValueInAnalog[#temp16IndexMTP].SclMinExt;
                                                   #ProcessInAna[#temp16IndexAnalog].SclMaxExt := #ProcessValueInAnalog[#temp16IndexMTP].SclMaxExt;
                                                   #ProcessInAna[#temp16IndexAnalog].UnitExt := #ProcessValueInAnalog[#temp16IndexMTP].UnitExt;
                                                   #ProcessInAna[#temp16IndexAnalog].Apply := #ProcessValueInAnalog[#temp16IndexMTP].Apply;
                                                   #ProcessInAna[#temp16IndexAnalog].ApplyEn := #ProcessValueInAnalog[#temp16IndexMTP].ApplyEn;
                                               END_IF;
                                               #temp16IndexAnalog := #temp16IndexAnalog + 1;
                                           END_REGION
                                       #TYPE_DIGITAL:
                                           REGION Digital
                                               //Bit Masking funtionality for calculate the used Digital parameter and Position of the Parameter name in the HMI Text List 
                                               #ProcessInValueType.IndexDigital := #ProcessInValueType.IndexDigital OR SHL(IN := #temp32TempDword1, N := INT_TO_UINT(#temp16IndexOfDefinitionProcessIn));
                                               #ProcessInValueType.NameIndexDigital := #ProcessInValueType.NameIndexDigital OR SHL(IN := #temp32TempDword1, N := INT_TO_UINT(#temp16IndexOfDefinition));
                                               IF ((#temp16IndexIO >= #PROCESS_VALUES_IN_MIN) AND (#temp16IndexIO <= #PROCESS_VALUES_IN_DIGITAL_MAX)) THEN
                                                   //WinCC Parameter View Faceplate logic
                                                   #ProcessInDint[#temp16IndexDigital].WQC := #ProcessValueInDigital[#temp16IndexMTP].WQC;
                                                   #ProcessInDint[#temp16IndexDigital].OSLevel := #ProcessValueInDigital[#temp16IndexMTP].OSLevel;
                                                   #ProcessInDint[#temp16IndexDigital].V := #ProcessValueInDigital[#temp16IndexMTP].V;
                                                   #ProcessInDint[#temp16IndexDigital].VQC := #ProcessValueInDigital[#temp16IndexMTP].VQC;
                                                   #ProcessInDint[#temp16IndexDigital].SclMinCur := #ProcessValueInDigital[#temp16IndexMTP].SclMinCur;
                                                   #ProcessInDint[#temp16IndexDigital].SclMaxCur := #ProcessValueInDigital[#temp16IndexMTP].SclMaxCur;
                                                   #ProcessInDint[#temp16IndexDigital].UnitCur := #ProcessValueInDigital[#temp16IndexMTP].UnitCur;
                                                   #ProcessInDint[#temp16IndexDigital].SclMinExt := #ProcessValueInDigital[#temp16IndexMTP].SclMinExt;
                                                   #ProcessInDint[#temp16IndexDigital].SclMaxExt := #ProcessValueInDigital[#temp16IndexMTP].SclMaxExt;
                                                   #ProcessInDint[#temp16IndexDigital].UnitExt := #ProcessValueInDigital[#temp16IndexMTP].UnitExt;
                                                   #ProcessInDint[#temp16IndexDigital].Apply := #ProcessValueInDigital[#temp16IndexMTP].Apply;
                                                   #ProcessInDint[#temp16IndexDigital].ApplyEn := #ProcessValueInDigital[#temp16IndexMTP].ApplyEn;
                                               END_IF;
                                               #temp16IndexDigital := #temp16IndexDigital + 1;
                                           END_REGION
                                       #TYPE_BINARY:
                                           REGION Binary
                                               //Bit Masking funtionality for calculate the used Binary parameter and Position of the Parameter name in the HMI Text List 
                                               #ProcessInValueType.IndexBinary := #ProcessInValueType.IndexBinary OR SHL(IN := #temp32TempDword1, N := INT_TO_UINT(#temp16IndexOfDefinitionProcessIn));
                                               #ProcessInValueType.NameIndexBinary := #ProcessInValueType.NameIndexBinary OR SHL(IN := #temp32TempDword1, N := INT_TO_UINT(#temp16IndexOfDefinition));
                                               IF ((#temp16IndexIO >= #PROCESS_VALUES_IN_MIN) AND (#temp16IndexIO <= #PROCESS_VALUES_IN_BINARY_MAX)) THEN
                                                   //WinCC Parameter View Faceplate logic
                                                   #ProcessInBin[#temp16IndexBinary].WQC := #ProcessValueInBinary[#temp16IndexMTP].WQC;
                                                   #ProcessInBin[#temp16IndexBinary].V := #ProcessValueInBinary[#temp16IndexMTP].V;
                                                   #ProcessInBin[#temp16IndexBinary].VQC := #ProcessValueInBinary[#temp16IndexMTP].VQC;
                                                   #ProcessInBin[#temp16IndexBinary].VState0 := #ProcessValueInBinary[#temp16IndexMTP].VState0;
                                                   #ProcessInBin[#temp16IndexBinary].VState1 := #ProcessValueInBinary[#temp16IndexMTP].VState1;
                                               END_IF;
                                               #temp16IndexBinary := #temp16IndexBinary + 1;
                                           END_REGION
                                       #TYPE_STRING:
                                           REGION String
                                               //Bit Masking funtionality for calculate the used String parameter and Position of the Parameter name in the HMI Text List 
                                               #ProcessInValueType.IndexString := #ProcessInValueType.IndexString OR SHL(IN := #temp32TempDword1, N := INT_TO_UINT(#temp16IndexOfDefinitionProcessIn));
                                               #ProcessInValueType.NameIndexString := #ProcessInValueType.NameIndexString OR SHL(IN := #temp32TempDword1, N := INT_TO_UINT(#temp16IndexOfDefinition));
                                               IF ((#temp16IndexIO >= #PROCESS_VALUES_IN_MIN) AND (#temp16IndexIO <= #PROCESS_VALUES_IN_STRING_MAX)) THEN
                                                   //WinCC Parameter View Faceplate logic
                                                   #ProcessInString[#temp16IndexString].WQC := #ProcessValueInString[#temp16IndexMTP].WQC;
                                                   #ProcessInString[#temp16IndexString].V := #ProcessValueInString[#temp16IndexMTP].V;
                                                   #ProcessInString[#temp16IndexString].VQC := #ProcessValueInString[#temp16IndexMTP].VQC;
                                               END_IF;
                                               #temp16IndexString := #temp16IndexString + 1;
                                           END_REGION
                                   END_CASE;
                               END_IF;
                           END_IF;
                           #temp16IndexOfDefinitionProcessIn := #temp16IndexOfDefinitionProcessIn + 1;
                       END_IF;
                   END_FOR;
               END_IF;
           END_IF;
       END_REGION

       REGION Process Out Values

           REGION Get Start and End index details of the Current /Prepared procedure
               //Current/Prepared procedure selection for parameter display in the faceplate
               //#stat32PrecedureProcessOutMap := -1;
               IF NOT (#ProcessOutValueType.ProcedureReqCurInd) THEN
                   #stat32PrecedureProcessOutMap := #tempSetup.procedure.procedure[#stat16ProceCurIndex].ProcedureProcessOutMap[0];
               ELSIF (#ProcessOutValueType.ProcedureReqCurInd) THEN
                   #stat32PrecedureProcessOutMap := #tempSetup.procedure.procedure[#stat16ProceReqIndex].ProcedureProcessOutMap[0];
               END_IF;
           END_REGION
           //Initialize the used variable values          
           #temp32TempDword1 := 16#1;
           #temp16IndexAnalog := 16#0;
           #temp16IndexDigital := 16#0;
           #temp16IndexBinary := 16#0;
           #temp16IndexString := 16#0;
           //Initialize the Process Out Value index and Name index while changing of Procedure and changing of screen selection b/w Prepared and Current procedure
           IF ((#statLasProcedureCur <> #ProcedureCur) OR (#statLasProcedureReq <> #ProcedureReq) OR (#StatLastProceselProcessOut <> #ProcessOutValueType.ProcedureReqCurInd)
               OR (((#ProcedureCur = 16#0) AND NOT #ProcessOutValueType.ProcedureReqCurInd) OR ((#ProcedureReq = 16#0) AND #ProcessOutValueType.ProcedureReqCurInd))) THEN
               #ProcessOutValueType.IndexAnalog := 16#0;
               #ProcessOutValueType.NameIndexAnalog := 16#0;
               #ProcessOutValueType.IndexDigital := 16#0;
               #ProcessOutValueType.NameIndexDigital := 16#0;
               #ProcessOutValueType.IndexBinary := 16#0;
               #ProcessOutValueType.NameIndexBinary := 16#0;
               #ProcessOutValueType.IndexString := 16#0;
               #ProcessOutValueType.NameIndexString := 16#0;
           END_IF;
           //Used/Mapped parameter count with individual parameter type will written from the Tool
           #statTotalProcessOutValues := #MAPPED_PROCESS_OUT_ANALOG + #MAPPED_PROCESS_OUT_DIGITAL + #MAPPED_PROCESS_OUT_BINARY + #MAPPED_PROCESS_OUT_STRING - 1;
           IF (((#ProcedureCur <> 16#0) AND NOT #ProcessOutValueType.ProcedureReqCurInd) OR ((#ProcedureReq <> 16#0) AND #ProcessOutValueType.ProcedureReqCurInd)) THEN
               IF ((#statTotalProcessOutValues >= 0) AND (#statTotalProcessOutValues <= #PROCESS_VALUES_OUT_MAX)) THEN
                   #temp16IndexOfDefinitionProcessOut := 16#0;
                   FOR #temp16IndexOfDefinition := #PROCESS_VALUES_OUT_MIN TO #statTotalProcessOutValues BY 1 DO
                       #temp16ParameterCMAddress := BYTE_TO_INT(#tempSetup.processValueOutData.definition[#temp16IndexOfDefinition].controlModule);
                       #temp16ParameterType := #tempSetup.processValueOutData.definition[#temp16IndexOfDefinition].type;
                       #temp16IndexMTP := #tempSetup.processValueOutData.definition[#temp16IndexOfDefinition].indexMTP;
                       #tempUsed := #tempSetup.processValueOutData.used;
                       // Find the procedure information assigned with the processOut values
                       IF (((#stat32PrecedureProcessOutMap AND SHL(IN := #temp32TempDword1, N := INT_TO_UINT(#temp16IndexOfDefinition))) <> 0) = TRUE) THEN
                           #temp16IndexIO := #tempSetup.processValueOutData.definition[#temp16IndexOfDefinition].indexIO;

                           IF (#temp16ParameterCMAddress <> 255) AND (#temp16ParameterCMAddress >= #NUMBER_OF_CONTROLMODULES_MIN) AND (#temp16ParameterCMAddress <= #NUMBER_OF_CONTROLMODULES)
                               AND (#temp16ParameterType >= #TYPE_NONE) AND (#temp16ParameterType <= #TYPE_STRING) THEN
                               #temp16TempInt1 := #temp16ParameterCMAddress / 32;    //DWORD - Adress
                               #temp16TempInt2 := #temp16ParameterCMAddress MOD 32;  //Bit - Adress
                               //If parameter is forced (FRC) --> Parameter is used
                               IF (((#tempUsed[#temp16TempInt1] AND SHL(IN := #temp32TempDword1, N := INT_TO_UINT(#temp16TempInt2))) <> 0) = TRUE) THEN
                                   CASE #temp16ParameterType OF
                                       #TYPE_ANALOG:
                                           REGION Analog
                                               //Bit Masking funtionality for calculate the used Analog parameter and Position of the Parameter name in the HMI Text List                                         
                                               #ProcessOutValueType.IndexAnalog := #ProcessOutValueType.IndexAnalog OR SHL(IN := #temp32TempDword1, N := INT_TO_UINT(#temp16IndexOfDefinitionProcessOut));
                                               #ProcessOutValueType.NameIndexAnalog := #ProcessOutValueType.NameIndexAnalog OR SHL(IN := #temp32TempDword1, N := INT_TO_UINT(#temp16IndexOfDefinition));
                                               IF ((#temp16IndexIO >= #PROCESS_VALUES_OUT_MIN) AND (#temp16IndexIO <= #PROCESS_VALUES_OUT_ANALOG_MAX)) THEN
                                                   //WinCC Parameter View Faceplate logic
                                                   #ProcessOutAna[#temp16IndexAnalog].WQC := #ProcessValueOutAnalog[#temp16IndexMTP].WQC;
                                                   #ProcessOutAna[#temp16IndexAnalog].V := #ProcessValueOutAnalog[#temp16IndexMTP].V;
                                                   #ProcessOutAna[#temp16IndexAnalog].VSclMin := #ProcessValueOutAnalog[#temp16IndexMTP].VSclMin;
                                                   #ProcessOutAna[#temp16IndexAnalog].VSclMax := #ProcessValueOutAnalog[#temp16IndexMTP].VSclMax;
                                                   #ProcessOutAna[#temp16IndexAnalog].VUnit := #ProcessValueOutAnalog[#temp16IndexMTP].VUnit;
                                               END_IF;
                                               #temp16IndexAnalog := #temp16IndexAnalog + 1;
                                           END_REGION
                                       #TYPE_DIGITAL:
                                           REGION Digital
                                               //Bit Masking funtionality for calculate the used Digital parameter and Position of the Parameter name in the HMI Text List                                         
                                               #ProcessOutValueType.IndexDigital := #ProcessOutValueType.IndexDigital OR SHL(IN := #temp32TempDword1, N := INT_TO_UINT(#temp16IndexOfDefinitionProcessOut));
                                               #ProcessOutValueType.NameIndexDigital := #ProcessOutValueType.NameIndexDigital OR SHL(IN := #temp32TempDword1, N := INT_TO_UINT(#temp16IndexOfDefinition));
                                               IF ((#temp16IndexIO >= #PROCESS_VALUES_OUT_MIN) AND (#temp16IndexIO <= #PROCESS_VALUES_OUT_DIGITAL_MAX)) THEN
                                                   //WinCC Parameter View Faceplate logic
                                                   #ProcessOutDint[#temp16IndexDigital].WQC := #ProcessValueOutDigital[#temp16IndexMTP].WQC;
                                                   #ProcessOutDint[#temp16IndexDigital].V := #ProcessValueOutDigital[#temp16IndexMTP].V;
                                                   #ProcessOutDint[#temp16IndexDigital].VSclMin := #ProcessValueOutDigital[#temp16IndexMTP].VSclMin;
                                                   #ProcessOutDint[#temp16IndexDigital].VSclMax := #ProcessValueOutDigital[#temp16IndexMTP].VSclMax;
                                                   #ProcessOutDint[#temp16IndexDigital].VUnit := #ProcessValueOutDigital[#temp16IndexMTP].VUnit;
                                               END_IF;
                                               #temp16IndexDigital := #temp16IndexDigital + 1;
                                           END_REGION
                                       #TYPE_BINARY:
                                           REGION Binary
                                               //Bit Masking funtionality for calculate the used Binary parameter and Position of the Parameter name in the HMI Text List 
                                               #ProcessOutValueType.IndexBinary := #ProcessOutValueType.IndexBinary OR SHL(IN := #temp32TempDword1, N := INT_TO_UINT(#temp16IndexOfDefinitionProcessOut));
                                               #ProcessOutValueType.NameIndexBinary := #ProcessOutValueType.NameIndexBinary OR SHL(IN := #temp32TempDword1, N := INT_TO_UINT(#temp16IndexOfDefinition));
                                               IF ((#temp16IndexIO >= #PROCESS_VALUES_OUT_MIN) AND (#temp16IndexIO <= #PROCESS_VALUES_OUT_BINARY_MAX)) THEN
                                                   //WinCC Parameter View Faceplate logic
                                                   #ProcessOutBin[#temp16IndexBinary].WQC := #ProcessValueOutBinary[#temp16IndexMTP].WQC;
                                                   #ProcessOutBin[#temp16IndexBinary].V := #ProcessValueOutBinary[#temp16IndexMTP].V;
                                                   #ProcessOutBin[#temp16IndexBinary].VState0 := #ProcessValueOutBinary[#temp16IndexMTP].VState0;
                                                   #ProcessOutBin[#temp16IndexBinary].VState1 := #ProcessValueOutBinary[#temp16IndexMTP].VState1;
                                               END_IF;
                                               #temp16IndexBinary := #temp16IndexBinary + 1;
                                           END_REGION
                                       #TYPE_STRING:
                                           REGION String
                                               //Bit Masking funtionality for calculate the used String parameter and Position of the Parameter name in the HMI Text List 
                                               #ProcessOutValueType.IndexString := #ProcessOutValueType.IndexString OR SHL(IN := #temp32TempDword1, N := INT_TO_UINT(#temp16IndexOfDefinitionProcessOut));
                                               #ProcessOutValueType.NameIndexString := #ProcessOutValueType.NameIndexString OR SHL(IN := #temp32TempDword1, N := INT_TO_UINT(#temp16IndexOfDefinition));
                                               IF ((#temp16IndexIO >= #PROCESS_VALUES_OUT_MIN) AND (#temp16IndexIO <= #PROCESS_VALUES_OUT_STRING_MAX)) THEN
                                                   //WinCC Parameter View Faceplate logic
                                                   #ProcessOutString[#temp16IndexString].WQC := #ProcessValueOutString[#temp16IndexMTP].WQC;
                                                   #ProcessOutString[#temp16IndexString].Text := #ProcessValueOutString[#temp16IndexMTP].Text;
                                               END_IF;
                                               #temp16IndexString := #temp16IndexString + 1;
                                           END_REGION
                                   END_CASE;
                               END_IF;
                           END_IF;
                           #temp16IndexOfDefinitionProcessOut := #temp16IndexOfDefinitionProcessOut + 1;
                       END_IF;
                   END_FOR;
               END_IF;
           END_IF;
       END_REGION

       REGION Report Values

           REGION Get Start and End index details of the Current /Prepared procedure
               //Current/Prepared procedure selection for parameter display in the faceplate
              // #stat32PrecedureReportMap := -1;
               IF NOT (#ReportValueType.ProcedureReqCurInd) THEN
                   #stat32PrecedureReportMap := #tempSetup.procedure.procedure[#stat16ProceCurIndex].ProcedureReportMap[0];
               ELSIF (#ReportValueType.ProcedureReqCurInd) THEN
                   #stat32PrecedureReportMap := #tempSetup.procedure.procedure[#stat16ProceReqIndex].ProcedureReportMap[0];
               END_IF;
           END_REGION
           //Initialize the used variable values        
           #temp32TempDword1 := 16#1;
           #temp16IndexAnalog := 16#0;
           #temp16IndexDigital := 16#0;
           #temp16IndexBinary := 16#0;
           #temp16IndexString := 16#0;
           //Initialize the Process Out Value index and Name index while changing of Procedure and changing of screen selection b/w Prepared and Current procedure
           IF ((#statLasProcedureCur <> #ProcedureCur) OR (#statLasProcedureReq <> #ProcedureReq) OR (#StatLastProceselReport <> #ReportValueType.ProcedureReqCurInd)
               OR (((#ProcedureCur = 16#0) AND NOT #ReportValueType.ProcedureReqCurInd) OR ((#ProcedureReq = 16#0) AND #ReportValueType.ProcedureReqCurInd))) THEN
               #ReportValueType.IndexAnalog := 16#0;
               #ReportValueType.NameIndexAnalog := 16#0;
               #ReportValueType.IndexDigital := 16#0;
               #ReportValueType.NameIndexDigital := 16#0;
               #ReportValueType.IndexBinary := 16#0;
               #ReportValueType.NameIndexBinary := 16#0;
               #ReportValueType.IndexString := 16#0;
               #ReportValueType.NameIndexString := 16#0;
           END_IF;
           //Used/Mapped parameter count with individual parameter type will written from the Tool
           #statTotalReportValues := #MAPPED_REPORT_ANALOG + #MAPPED_REPORT_DIGITAL + #MAPPED_REPORT_BINARY + #MAPPED_REPORT_STRING - 1;
           IF (((#ProcedureCur <> 16#0) AND NOT #ReportValueType.ProcedureReqCurInd) OR ((#ProcedureReq <> 16#0) AND #ReportValueType.ProcedureReqCurInd)) THEN
               IF ((#statTotalReportValues >= 0) AND (#statTotalReportValues <= #REPORT_VALUES_MAX)) THEN
                   #temp16IndexOfDefinitionReport := 16#0;
                   FOR #temp16IndexOfDefinition := #REPORT_VALUES_MIN TO #statTotalReportValues BY 1 DO
                       #temp16ParameterCMAddress := BYTE_TO_INT(#tempSetup.reportValueData.definition[#temp16IndexOfDefinition].controlModule);
                       #temp16ParameterType := #tempSetup.reportValueData.definition[#temp16IndexOfDefinition].type;
                       #temp16IndexMTP := #tempSetup.reportValueData.definition[#temp16IndexOfDefinition].indexMTP;
                       #tempUsed := #tempSetup.reportValueData.used;
                       // Find the procedure information assigned with the report values
                       IF (((#stat32PrecedureReportMap AND SHL(IN := #temp32TempDword1, N := INT_TO_UINT(#temp16IndexOfDefinition))) <> 0) = TRUE) THEN
                           #temp16IndexIO := #tempSetup.reportValueData.definition[#temp16IndexOfDefinition].indexIO;

                           IF (#temp16ParameterCMAddress <> 255) AND (#temp16ParameterCMAddress >= #NUMBER_OF_CONTROLMODULES_MIN) AND (#temp16ParameterCMAddress <= #NUMBER_OF_CONTROLMODULES)
                               AND (#temp16ParameterType >= #TYPE_NONE) AND (#temp16ParameterType <= #TYPE_STRING) THEN
                               #temp16TempInt1 := #temp16ParameterCMAddress / 32;    //DWORD - Adress
                               #temp16TempInt2 := #temp16ParameterCMAddress MOD 32;  //Bit - Adress
                               //If parameter is forced (FRC) --> Parameter is used
                               IF (((#tempUsed[#temp16TempInt1] AND SHL(IN := #temp32TempDword1, N := INT_TO_UINT(#temp16TempInt2))) <> 0) = TRUE) THEN
                                   CASE #temp16ParameterType OF
                                       #TYPE_ANALOG:
                                           REGION Analog
                                               //Bit Masking funtionality for calculate the used Analog parameter and Position of the Parameter name in the HMI Text List 
                                               #ReportValueType.IndexAnalog := #ReportValueType.IndexAnalog OR SHL(IN := #temp32TempDword1, N := INT_TO_UINT(#temp16IndexOfDefinitionReport));
                                               #ReportValueType.NameIndexAnalog := #ReportValueType.NameIndexAnalog OR SHL(IN := #temp32TempDword1, N := INT_TO_UINT(#temp16IndexOfDefinition));
                                               IF ((#temp16IndexIO >= #REPORT_VALUES_MIN) AND (#temp16IndexIO <= #REPORT_VALUES_ANALOG_MAX)) THEN
                                                   //WinCC Parameter View Faceplate logic
                                                   #ReportAna[#temp16IndexAnalog].WQC := #ReportValueAnalog[#temp16IndexMTP].WQC;
                                                   #ReportAna[#temp16IndexAnalog].V := #ReportValueAnalog[#temp16IndexMTP].V;
                                                   #ReportAna[#temp16IndexAnalog].VSclMin := #ReportValueAnalog[#temp16IndexMTP].VSclMin;
                                                   #ReportAna[#temp16IndexAnalog].VSclMax := #ReportValueAnalog[#temp16IndexMTP].VSclMax;
                                                   #ReportAna[#temp16IndexAnalog].VUnit := #ReportValueAnalog[#temp16IndexMTP].VUnit;
                                                   #ReportAna[#temp16IndexAnalog].MissedValue := #ReportValueAnalog[#temp16IndexMTP].MissedValue;
                                               END_IF;
                                               #temp16IndexAnalog := #temp16IndexAnalog + 1;
                                           END_REGION
                                       #TYPE_DIGITAL:
                                           REGION Digital
                                               //Bit Masking funtionality for calculate the used Digital parameter and Position of the Parameter name in the HMI Text List 
                                               #ReportValueType.IndexDigital := #ReportValueType.IndexDigital OR SHL(IN := #temp32TempDword1, N := INT_TO_UINT(#temp16IndexOfDefinitionReport));
                                               #ReportValueType.NameIndexDigital := #ReportValueType.NameIndexDigital OR SHL(IN := #temp32TempDword1, N := INT_TO_UINT(#temp16IndexOfDefinition));
                                               IF ((#temp16IndexIO >= #REPORT_VALUES_MIN) AND (#temp16IndexIO <= #REPORT_VALUES_DIGITAL_MAX)) THEN
                                                   //WinCC Parameter View Faceplate logic
                                                   #ReportDint[#temp16IndexDigital].WQC := #ReportValueDigital[#temp16IndexMTP].WQC;
                                                   #ReportDint[#temp16IndexDigital].V := #ReportValueDigital[#temp16IndexMTP].V;
                                                   #ReportDint[#temp16IndexDigital].VSclMin := #ReportValueDigital[#temp16IndexMTP].VSclMin;
                                                   #ReportDint[#temp16IndexDigital].VSclMax := #ReportValueDigital[#temp16IndexMTP].VSclMax;
                                                   #ReportDint[#temp16IndexDigital].VUnit := #ReportValueDigital[#temp16IndexMTP].VUnit;
                                                   #ReportDint[#temp16IndexDigital].MissedValue := #ReportValueDigital[#temp16IndexMTP].MissedValue;
                                               END_IF;
                                               #temp16IndexDigital := #temp16IndexDigital + 1;
                                           END_REGION
                                       #TYPE_BINARY:
                                           REGION Binary
                                               //Bit Masking funtionality for calculate the used Binary parameter and Position of the Parameter name in the HMI Text List 
                                               #ReportValueType.IndexBinary := #ReportValueType.IndexBinary OR SHL(IN := #temp32TempDword1, N := INT_TO_UINT(#temp16IndexOfDefinitionReport));
                                               #ReportValueType.NameIndexBinary := #ReportValueType.NameIndexBinary OR SHL(IN := #temp32TempDword1, N := INT_TO_UINT(#temp16IndexOfDefinition));
                                               IF ((#temp16IndexIO >= #REPORT_VALUES_MIN) AND (#temp16IndexIO <= #REPORT_VALUES_BINARY_MAX)) THEN
                                                   //WinCC Parameter View Faceplate logic
                                                   #ReportBin[#temp16IndexBinary].WQC := #ReportValueBinary[#temp16IndexMTP].WQC;
                                                   #ReportBin[#temp16IndexBinary].V := #ReportValueBinary[#temp16IndexMTP].V;
                                                   #ReportBin[#temp16IndexBinary].VState0 := #ReportValueBinary[#temp16IndexMTP].VState0;
                                                   #ReportBin[#temp16IndexBinary].VState1 := #ReportValueBinary[#temp16IndexMTP].VState1;
                                                   #ReportBin[#temp16IndexBinary].MissedValue := #ReportValueBinary[#temp16IndexMTP].MissedValue;
                                               END_IF;
                                               #temp16IndexBinary := #temp16IndexBinary + 1;
                                           END_REGION
                                       #TYPE_STRING:
                                           REGION String
                                               //Bit Masking funtionality for calculate the used String parameter and Position of the Parameter name in the HMI Text List 
                                               #ReportValueType.IndexString := #ReportValueType.IndexString OR SHL(IN := #temp32TempDword1, N := INT_TO_UINT(#temp16IndexOfDefinitionReport));
                                               #ReportValueType.NameIndexString := #ReportValueType.NameIndexString OR SHL(IN := #temp32TempDword1, N := INT_TO_UINT(#temp16IndexOfDefinition));
                                               IF ((#temp16IndexIO >= #REPORT_VALUES_MIN) AND (#temp16IndexIO <= #REPORT_VALUES_STRING_MAX)) THEN

                                                   //WinCC Parameter View Faceplate logic
                                                   #ReportString[#temp16IndexString].WQC := #ReportValueString[#temp16IndexMTP].WQC;
                                                   #ReportString[#temp16IndexString].Text := #ReportValueString[#temp16IndexMTP].Text;
                                                   #ReportString[#temp16IndexString].MissedValue := #ReportValueString[#temp16IndexMTP].MissedValue;
                                               END_IF;
                                               #temp16IndexString := #temp16IndexString + 1;
                                           END_REGION
                                   END_CASE;
                               END_IF;
                           END_IF;
                           #temp16IndexOfDefinitionReport := #temp16IndexOfDefinitionReport + 1;
                       END_IF;
                   END_FOR;
               END_IF;
           END_IF;
       END_REGION  

       //Move last valid value 
       #statLasProcedureCur := #ProcedureCur;
       #statLasProcedureReq := #ProcedureReq;
       #statLastReqProcedSelected := #ProcedureParaType.ProcedureReqCurInd;
       #StatLastProceselProcessIn := #ProcessInValueType.ProcedureReqCurInd;
       #StatLastProceselProcessOut := #ProcessOutValueType.ProcedureReqCurInd;
       #StatLastProceselReport := #ReportValueType.ProcedureReqCurInd;
END_FUNCTION_BLOCK
